// TIA Portal V20 export
VAR_GLOBAL   // PLC tag table "Hauptvariablen"
   DE_Bedienerkonsole_Taste_K0_leer AT %I20.0 : Bool;   // +SK2-458K2 Bedienerkonsole Taste K0 leer
   DE_Bedienerkonsole_Taste_K1_Stopp AT %I20.1 : Bool;   // +SK2-458K2 Bedienerkonsole Taste K1 Stopp
   DE_Bedienerkonsole_Taste_K2_ACK AT %I20.2 : Bool;   // +SK2-458K2 Bedienerkonsole Taste K2 ACK
   DE_Bedienerkonsole_Taste_K3_Start AT %I20.3 : Bool;   // +SK2-458K2 Bedienerkonsole Taste K3 Start
   DE_Bedienerkonsole_Taste_K4_Verwaltung AT %I20.4 : Bool;   // +SK2-458K2 Bedienerkonsole Taste K4 leer
   DE_Bedienerkonsole_Taste_K5_Richten AT %I20.5 : Bool;   // +SK2-458K2 Bedienerkonsole Taste K5 Betriebsart Richten
   DE_Bedienerkonsole_Taste_K6_Manuell AT %I20.6 : Bool;   // +SK2-458K2 Bedienerkonsole Taste K6 Betriebsart Manuell
   "DE_Bedienerkonsole Taste_K7_Automatik" AT %I20.7 : Bool;   // +SK2-458K2 Bedienerkonsole Taste K7 Betriebsart Automatik
   DE_Bedienerkonsole_DE_0 AT %I21.0 : Bool;   // +SK2-458K2 Bedienerkonsole Digital Eingang 0
   DE_Bedienerkonsole_DE_1 AT %I21.1 : Bool;   // +SK2-458K2 Bedienerkonsole Digital Eingang 1
   DE_Bedienerkonsole_DE_2 AT %I21.2 : Bool;   // +SK2-458K2 Bedienerkonsole Digital Eingang 2
   DE_Bedienerkonsole_DE_3 AT %I21.3 : Bool;   // +SK2-458K2 Bedienerkonsole Digital Eingang 3
   DE_Bedienerkonsole_DE_4 AT %I21.4 : Bool;   // +SK2-458K2 Bedienerkonsole Digital Eingang 4
   DE_Bedienerkonsole_DE_5 AT %I21.5 : Bool;   // +SK2-458K2 Bedienerkonsole Digital Eingang 5
   DE_Bedienerkonsole_DE_6 AT %I21.6 : Bool;   // +SK2-458K2 Bedienerkonsole Digital Eingang 6
   DE_Bedienerkonsole_DE_7 AT %I21.7 : Bool;   // +SK2-458K2 Bedienerkonsole Digital Eingang 7
END_VAR
